(* IEC 61131-3 sources: codesys-to-s7/tests/corpus/C2S7-NAME-KEYWORD/neg, 1 file *)

(* ---- input.st ---- *)
FUNCTION_BLOCK FB_Case
VAR
    xBegin : INT;
END_VAR
xBegin := 1;
END_FUNCTION_BLOCK
